// TIA Portal V20 export
// export: Created 2026-10-11T05:22:23.299998Z, ExportSetting WithDefaults, DisplayName Totally Integrated Automation Portal, DisplayVersion V20, DisplayName TIA Portal Openness, DisplayVersion V20, DisplayName TIA Portal Teamcenter Gateway, DisplayVersion V20, DisplayName TIA Portal Version Control Interface, DisplayVersion V20, DisplayName SINAMICS Startdrive Advanced, DisplayVersion V20 SP1 Update 2, DisplayName SINAMICS Startdrive G110M, G120, G120C, G120D, G120P, G115D, DisplayVersion V20 SP1 Update 2, DisplayName SINAMICS Startdrive G130, G150, S120, S150, SINAMICS MV, G220, S200, S210, DisplayVersion V20 SP1 Update 2, DisplayName STEP 7 Professional, DisplayVersion V20, DisplayName STEP 7 Safety, DisplayVersion V20, DisplayName WinCC Basic/Comfort/Advanced, DisplayVersion V20, DisplayName WinCC Professional, DisplayVersion V20, DisplayName WinCC Unified, DisplayVersion V20
FUNCTION "FRK_Diagnostic" : Void   // FC7, SCL
{ S7_Optimized_Access := 'TRUE' }
VERSION : 0.1
// stored: AutoNumber true, IsIECCheckEnabled false, SetENOAutomatically false, UDAEnableTagReadback false
   VAR_INPUT
      ReasonCode : DInt;
      Description : WString;
      Severity : DInt;
   END_VAR
   VAR_IN_OUT
      Status : "ST_ModuleStatus";
   END_VAR
   VAR_TEMP
      Stamp : DTL;
      ResultCode : Int;
   END_VAR
BEGIN

   #Status.Diagnostic.ReasonCode := #ReasonCode;
   #Status.Diagnostic.SourcePath := STRING_TO_WSTRING(#Status.Name);
   #Status.Diagnostic.Description := #Description;
   #Status.Diagnostic.IoTag := '';
   #Status.Diagnostic.IoAddress := '';
   #Status.Diagnostic.Severity := #Severity;
   #Status.Diagnostic.Category := 0;
   #ResultCode := RD_SYS_T(OUT => #Stamp);
   IF #ResultCode = 0 THEN
       #Status.Diagnostic.Since := DTL_TO_LDT(#Stamp);
   ELSE
       #Status.Diagnostic.Since := LDT#1970-01-01-00:00:00.000000000;
   END_IF;
   // UTC source alone is not proof of synchronization; quality stays false.
   #Status.Diagnostic.TimeSynchronized := FALSE;
END_FUNCTION
